FUNCTION_BLOCK FB_Alarmmanager
VAR_INPUT
END_VAR
VAR_OUTPUT
END_VAR
VAR
END_VAR

END_FUNCTION_BLOCK

(* stored: Version 1.1.0.1
   POU FB_Alarmmanager: Id {5f7f12f7-1acf-402f-9ddd-b7b0c33babe4}, SpecialFunc None *)
